// TIA Portal V21 export
// export: Created 2026-08-21T20:18:55.2081305Z, ExportSetting None, DisplayName Totally Integrated Automation Portal, DisplayVersion V21, DisplayName STEP 7 Professional, DisplayVersion V21, DisplayName STEP 7 Safety, DisplayVersion V21, DisplayName Tech WebApplication, DisplayVersion V21, DisplayName WinCC Basic/Comfort/Advanced, DisplayVersion V21, DisplayName WinCC Professional, DisplayVersion V21, DisplayName WinCC Unified, DisplayVersion V21
TYPE "UDT_MTP_BinMon"
TITLE = MTPDataObjectSUCLibrary/DataAssembly/BinView
   STRUCT
      VState0 { ExternalWritable := 'False'} : String[16] := '';   // Text replacement for false
      VState1 { ExternalWritable := 'False'} : String[16] := '';   // Text replacement for true
      OSLevel : Byte := 16#00;   // OSLevel variable
      WQC { ExternalWritable := 'False'} : Byte := 16#FF;   // Worst Quality Code variable
      V { ExternalWritable := 'False'} : Bool := FALSE;   // Value
      VFlutEn { ExternalWritable := 'False'} : Bool;   // Enable Fluttering Recognition1: enabled; 0: disabled
      VFlutTi : Real;   // Period of an active signal before it will be recognized as flutter-free, in s
      VFlutCnt : Int;   // Counts of the allowed fluttering signals in the defined period VFlutTi
      VFlutAct { ExternalWritable := 'False'} : Bool;   // Fluttering Signal recognized1: Fluttering Signal recognized 0: no Fluttering Signal recognized
   END_STRUCT;
END_TYPE
